// CFC twin of T_SafeSr_Tests: the same tests drawn as CFC diagrams, the way a TwinSAFE project is authored.
    FUNCTION_BLOCK T_SafeSr_Tests_CFC EXTENDS T_SafeCfcTestSuite
    VAR
    // Test_SetDominantLatch
    group_1 : T_SafeGroup;
    fb_1 : T_SafeSr(group := group_1);
END_VAR

Test_SetDominantLatch();

METHOD PRIVATE Test_SetDominantLatch
// note: this text did not pass the execution check against the stored diagram
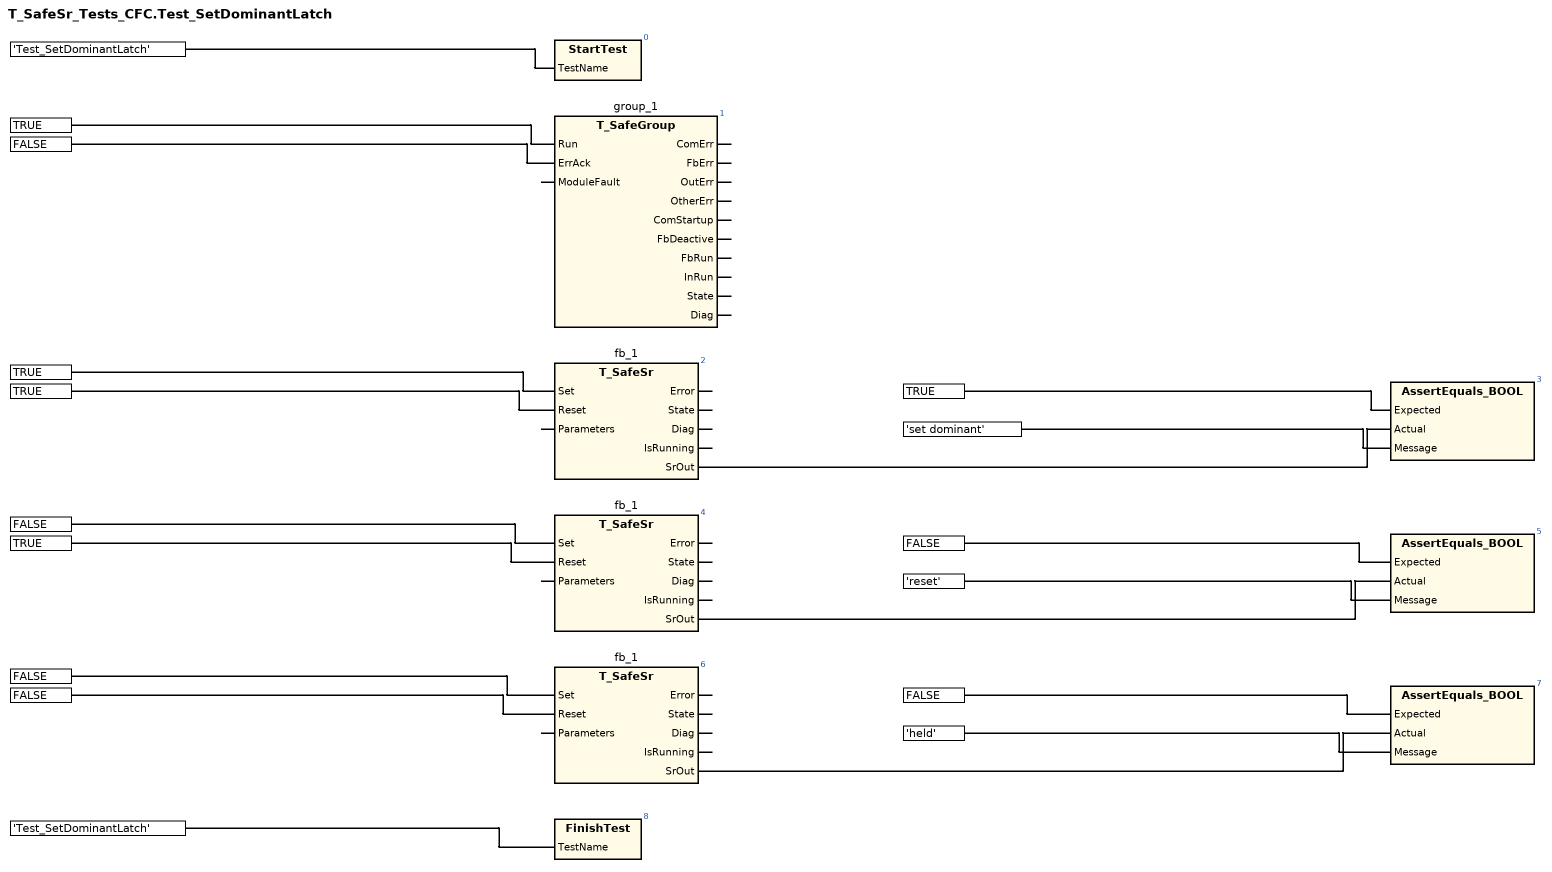
StartTest(TestName := 'Test_SetDominantLatch');
group_1(Run := TRUE, ErrAck := FALSE); // T_SafeGroup
fb_1(Set := TRUE, Reset := TRUE); // T_SafeSr
AssertEquals_BOOL(Expected := TRUE, Actual := fb_1.SrOut, Message := 'set dominant');
fb_1(Set := FALSE, Reset := TRUE); // T_SafeSr
AssertEquals_BOOL(Expected := FALSE, Actual := fb_1.SrOut, Message := 'reset');
fb_1(Set := FALSE, Reset := FALSE); // T_SafeSr
AssertEquals_BOOL(Expected := FALSE, Actual := fb_1.SrOut, Message := 'held');
FinishTest(TestName := 'Test_SetDominantLatch');
END_METHOD

END_FUNCTION_BLOCK

(* stored: Version 1.1.0.1, ProductVersion 3.1.4026.22
   POU T_SafeSr_Tests_CFC: Id {353c5686-7494-5336-bb25-8440a0f8bd1f}, SpecialFunc None
   Method Test_SetDominantLatch: Id {f7007b2e-affb-5b32-acbf-7d31d052b11f} *)
